(* IEC 61131-3 sources: POMIRTS_lab3/AS/Library_2/AsOpcUac, 3 files *)

(* ---- AsOpcUac.typ ---- *)
 TYPE
	UASecurityMsgMode :
	(												(* Message security modes *)
    	UASecurityMsgMode_BestAvailable 	:= 0,	(* Detects best available mode the server provides (may result in no security) 	*)
	  	UASecurityMsgMode_None          	:= 1,	(* No secure communication 														*)
	  	UASecurityMsgMode_Sign          	:= 2,	(* Messages are signed to verify peer authenticity 								*)
	  	UASecurityMsgMode_SignEncrypt   	:= 3	(* Messages are signed and encrypted 											*)
	);

  	UASecurityPolicy :
  	(												(* Security policies *)
    	UASecurityPolicy_BestAvailable  	:= 0,	(* Detects best available policy the server provides (may result in no security)	*)
    	UASecurityPolicy_None           	:= 1,	(* No secure communication (Allowed only for security mode = none)					*)
    	UASecurityPolicy_Basic128Rsa15  	:= 2,	(* RSA-PKCS-#1-V1.5-SHA1/RSA-PKCS-#1-V1.5/128-512 bit, HMAC-SHA1/AES-128-CBC/16bit	*)
    	UASecurityPolicy_Basic256       	:= 3,	(* RSA-PKCS-#1-OAEP-SHA1/RSA-OAEP/128-512 bit, HMAC-SHA1/AES-256-CBC/32bit			*)
    	UASecurityPolicy_Basic256Sha256   	:= 4	(* RSA-PKCS-#1-OAEP-SHA1/RSA-OAEP/256-512 bit, HMAC-SHA1/AES-256-CBC/32bit			*)
  	);

  	UATransportProfile :
  	(  												(* Transport profiles to select encoding and protocol *)
    	UATP_UATcp             				:= 1,	(* UA Binary over TCP								*)
    	UATP_WSHttpBinary      				:= 2,	(* Binary over HTTP			Not supported by B&R	*)
    	UATP_WSHttpXmlOrBinary 				:= 3,	(* XML/Binary over HTTP		Not supported by B&R	*)
    	UATP_WSHttpXml         				:= 4	(* XML over HTTP			Not supported by B&R	*)
  	);

 	UAUserIdentityTokenTtype :
 	(  												(* Authentication token type provided for logon *)
 		UAUITT_Anonymous					:= 0,	(* Logon anonymously					*)
 		UAUITT_Username						:= 1,	(* Logon with user name and password 	*)
 		UAUITT_x509							:= 2	(* Logon with user certificate			*)
 	);

	UAIdentifierType :
	(												(* Node identifier type *)
		UAIdentifierType_String 			:= 1,	(* String			*)
		UAIdentifierType_Numeric 			:= 2,	(* Numeric value	*)
		UAIdentifierType_GUID 				:= 3,	(* GUID				*)
		UAIdentifierType_Opaque				:= 4	(* ByteString		*)
	);

	UADeadbandType :
	(												(* Deadband type for monitored item sampling *)
		UADeadbandType_None 				:= 0,	(* No deadband, each value change is sampled						*)
		UADeadbandType_Absolute 			:= 1,	(* Absolute value to exceed from last sample to make new sample		*)
		UADeadbandType_Percent				:= 2	(* Percent of EURange to exceed from last sample to make new sample	*)
	);

	UANodeClass :
	(												(* Node classes defined through the OPC-UA standard *)
		UANodeClass_None 					:= 0,
		UANodeClass_Object					:= 1,
		UANodeClass_Variable 				:= 2,
		UANodeClass_Method					:= 4,
		UANodeClass_ObjectType				:= 8,
		UANodeClass_VariableType			:= 16,
		UANodeClass_ReferenceType			:= 32,
		UANodeClass_DataType				:= 64,
		UANodeClass_View					:= 128,
		UANodeClass_All						:= 255
	);

	UAAttributeId :
	(												(* Attributes defined through the OPC-UA standard *)
	  	UAAI_Default						:= 0,
		UAAI_NodeId							:= 1,
		UAAI_NodeClass						:= 2,
		UAAI_BrowseName						:= 3,
		UAAI_DisplayName					:= 4,
		UAAI_Description					:= 5,
		UAAI_WriteMask						:= 6,
		UAAI_UserWriteMask					:= 7,
		UAAI_IsAbstract						:= 8,
		UAAI_Symmetric						:= 9,
		UAAI_InverseName					:= 10,
		UAAI_ContainsNoLoops				:= 11,
		UAAI_EventNotifier					:= 12,
		UAAI_Value							:= 13,
		UAAI_DataType						:= 14,
		UAAI_ValueRank						:= 15,
		UAAI_ArrayDimensions				:= 16,
		UAAI_AccessLevel					:= 17,
		UAAI_UserAccessLevel				:= 18,
		UAAI_MinimumSamplingInterval		:= 19,
		UAAI_Historizing					:= 20,
		UAAI_Executable						:= 21,
		UAAI_UserExecutable					:= 22
	);

	UAConnectionStatus :
	(												(* Status of the underlying connection		*)
		UACS_Connected						:= 0,
		UACS_ConnectionError				:= 1,
		UACS_Shutdown						:= 2
	);

	UAServerState :
	(												(* State of the server read from Object.Server.ServerStatus.State	*)
		UASS_Running						:= 0,
		UASS_Failed							:= 1,
		UASS_NoConfiguration				:= 2,
		UASS_Suspended						:= 3,
		UASS_Shutdown						:= 4,
		UASS_Test							:= 5,
		UASS_CommunicationFault				:= 6,
		UASS_Unknown              			:= 7
	);

	UAVariantType :
	(												(* Kind of the variant data *)
		UAVariantType_Null					:= 0,	(* No data *)
		UAVariantType_Boolean				:= 1,	(* Data in element Boolean *)
		UAVariantType_SByte					:= 2,	(* Data in element SByte *)
		UAVariantType_Byte					:= 3,	(* Data in element Byte *)
		UAVariantType_Int16					:= 4,	(* Data in element Int16 *)
		UAVariantType_UInt16				:= 5,	(* Data in element UInt16 *)
		UAVariantType_Int32					:= 6,	(* Data in element Int32 *)
		UAVariantType_UInt32				:= 7,	(* Data in element UInt32 *)
		UAVariantType_Int64					:= 8,	(* Data in element Int64 *)
		UAVariantType_UInt64				:= 9,	(* Data in element UInt64 *)
		UAVariantType_Float					:= 10,	(* Data in element Float *)
		UAVariantType_Double				:= 11,	(* Data in element Double *)
		UAVariantType_String				:= 12,	(* Data in element String *)
		UAVariantType_DateTime				:= 13,	(* Data in element DateTime *)
		UAVariantType_Guid					:= 14,	(* Guid data in element String *)
		UAVariantType_ByteString			:= 15,	(* Byte string in element String *)
		UAVariantType_XmlElement			:= 16,	(* XML data in element String *)
		UAVariantType_NodeId				:= 17,	(* Data in element NodeId *)
		UAVariantType_ExpandedNodeId		:= 18,	(* Data in element ExpandedNodeId *)
		UAVariantType_StatusCode			:= 19,	(* Status code in element UInt32 *)
		UAVariantType_QualifiedName			:= 20,	(* Data in element QualifiedName *)
		UAVariantType_LocalizedText			:= 21	(* Data in element LocalizedText *)
	);

	UAArrayLength : DINT;							(* Arraylength of value attribute in AttributeRead and AttributeWrite services *)

	UANoOfElements : DINT;							(* Number of elements for arrays nested in structures *)

   	UAUserIdentityToken : STRUCT 					(* Identity token for authentication on an OPC-UA server *)
		UserIdentityTokenType	: UAUserIdentityTokenTtype;
		TokenParam1 			: STRING[255];
		TokenParam2				: STRING[255];
	END_STRUCT;

 	UASessionConnectInfo : STRUCT 					(* Session information and parameters *)
 	  	SessionName   			: STRING[255];
 	  	ApplicationName   		: STRING[255];
 	  	SecurityMsgMode   		: UASecurityMsgMode;
    	SecurityPolicy   		: UASecurityPolicy;
		CertificateStore		: STRING[255];
		ClientCertificateName	: STRING[255];
		ServerUri				: STRING[255];
		CheckServerCertificate	: BOOL;
    	TransportProfile 		: UATransportProfile;
    	UserIdentityToken		: UAUserIdentityToken;
		VendorSpecificParameter	: STRING[255];
    	SessionTimeout   		: TIME;
    	MonitorConnection		: TIME;
    	LocaleIDs				: ARRAY[0..4] OF STRING[6];
	END_STRUCT;

  	UANodeID : STRUCT 											(* Node identifier used to address nodes on the server		*)
		NamespaceIndex			: UINT;							(* Index of the namespace which contains the node			*)
		Identifier 				: STRING[255];					(* Node identifier according to the identifier types format *)
		IdentifierType			: UAIdentifierType; 			(* String, Numeric, GUID, ByteString						*)
	END_STRUCT;

	UAMonitoringSettings : STRUCT								(* Settings for data item monitoring						*)
		SamplingInterval		: TIME;							(* Time in ms 												*)
		DeadbandType			: UADeadbandType; 				(* Deadband type which applies to deadband value			*)
		Deadband				: REAL; 						(* Deadband value, semantics depending on DeadbandType 		*)
	END_STRUCT;

	UAMonitoringParameters : STRUCT								(* Settings for data item monitoring								*)
		SamplingInterval		: TIME;							(* Time in ms 														*)
		QueueSize				: UINT;							(* Size of the server sided queue to collect value changes			*)
		DiscardOldest			: BOOL;							(* True to discard oldest on queue overflow or newest otherwise		*)
		DeadbandType			: UADeadbandType; 				(* Deadband type which applies to deadband value					*)
		Deadband				: REAL; 						(* Deadband value, semantics depending on DeadbandType 				*)
	END_STRUCT;

	UALocalizedText : STRUCT									(* Localized text with locale identifer and text		*)
		Locale					: STRING[6];
		Text					: STRING[255];
	END_STRUCT;

	UANodeInfo : STRUCT											(* Node attribute values		*)
		AccessLevel 			: BYTE;
		ArrayDimension			: ARRAY[0..MAX_INDEX_ARRAYDIMENSION] OF UDINT;
		BrowseName				: STRING[255];
		ContainsNoLoops 		: BOOL;
		DataType				: UANodeID;
		Description				: UALocalizedText;
		DisplayName				: UALocalizedText;
		EventNotifier			: BYTE;
		Executable				: BOOL;
		Historizing				: BOOL;
		InverseName				: STRING[255];
		IsAbstract				: BOOL;
		MinimumSamplingInterval	: TIME;
		NodeClass				: UANodeClass;
		NodeID					: UANodeID;
		Symmetric				: BOOL;
		UserAccessLevel			: BYTE;
		UserExecutable			: BOOL;
		UserWriteMask			: UDINT;
		ValueRank				: DINT;
		WriteMask				: UDINT;
	END_STRUCT;

	UAIndexRange : STRUCT										(* Index range used for indexed access on arrays	*)
		StartIndex				: UINT;
		EndIndex 				: UINT;
	END_STRUCT;

	UANodeAdditionalInfo : STRUCT								(* Additional info for reading and writing node attributes	*)
		AttributeId				: UAAttributeId;
		IndexRangeCount			: UINT;
		IndexRange 				: ARRAY[0..MAX_INDEX_INDEXRANGE] OF UAIndexRange;
	END_STRUCT;

	UAMethodArgument : STRUCT						(* Method argument used to supply the input and receive the output argument values for method calls *)
		Name					: STRING[64];		(* Name of the method argument																		*)
		Value					: STRING[255];		(* Source/Destination variable name for the argument value											*)
	END_STRUCT;

	UAByteString : STRUCT							(* Byte string containing length and data	*)
		Length					: DINT;
		Data					: ARRAY[0..MAX_INDEX_BYTESTRING] OF USINT;
	END_STRUCT;

	UAExpandedNodeID : STRUCT 						(* Expanded node identfier type *)
		NodeId					: UANodeID;
		NamespaceUri			: STRING[255];
		ServerIndex				: UDINT;
	END_STRUCT;

	UAQualifiedName : STRUCT						(* Qualified name type *)
		NamespaceIndex			: UINT;
		Name					: STRING[255];
	END_STRUCT;

	UARelativePathElement : STRUCT					(* Relative path element used to build a relative path	*)
	    ReferenceTypeId			: UANodeID;
		IsInverse				: BOOL;
		IncludeSubTypes			: BOOL;
		TargetName				: UAQualifiedName;
	END_STRUCT;

	UARelativePath : STRUCT							(* Relative path used to translate and browse nodes	*)
	    NoOfElements			: DWORD;
		Elements				: ARRAY[0..MAX_INDEX_RELATIVEPATH] OF UARelativePathElement;
	END_STRUCT;

	UADataValue : STRUCT							(* Additional informations about data value *)
		Valid 					: BOOL;
		Reserved				: ARRAY[0..2]OF USINT;
		StatusCode				: UDINT;
		SourceTimestamp			: DATE_AND_TIME;
		ServerTimestamp			: DATE_AND_TIME;
	END_STRUCT;

	UAVariantData : STRUCT							(* Standard type for variant data *)
		VariantType				: UAVariantType;
		Boolean					: BOOL;
		SByte					: SINT;
		Byte					: USINT;
		Int16					: INT;
		UInt16					: UINT;
		Int32					: DINT;
		UInt32					: UDINT;
		Float					: REAL;
		Double					: LREAL;
		DateTime				: DATE_AND_TIME;
		String					: STRING[255];
		NodeId					: UANodeID;
		ExpandedNodeId			: UAExpandedNodeID;
		QualifiedName			: UAQualifiedName;
		LocalizedText			: UALocalizedText;
		DataValue				: UADataValue;
	END_STRUCT;

	UARange : STRUCT								(* Range for a value *)
		Low						: LREAL;
		High					: LREAL;
	END_STRUCT;

	UAEUInformation : STRUCT 						(* Information about the engineering units *)
		NamespaceUri			: STRING[255];
		UnitId					: DINT;
		DisplayName				: UALocalizedText;
		Description				: UALocalizedText;
	END_STRUCT;

	UATimeZoneData : STRUCT							(* Information about time zone	*)
		TimeOffset				: INT;				(* Offset in minutes from UTC	*)
		DaylightSaving			: BOOL;				(* Offset includes the DST		*)
	END_STRUCT;

	BrUaNodeId					: UANodeID;
	BrUaQualifiedName			: UAQualifiedName;
	BrUaLocalizedText			: UALocalizedText;
	BrUaByteString				: UAByteString;
	BrUaGuidString				: STRING[36];

	BrUaXmlElement : STRUCT
		Length					: DINT;
		Data					: STRING[65535];
	END_STRUCT;

	BrUaImageBMP : STRUCT
		Length					: DINT;
		Data					: ARRAY[0..6291455] OF USINT;
	END_STRUCT;
	BrUaImageGIF : STRUCT
		Length					: DINT;
		Data					: ARRAY[0..524287] OF USINT;
	END_STRUCT;
	BrUaImageJPG : STRUCT
		Length					: DINT;
		Data					: ARRAY[0..1048575] OF USINT;
	END_STRUCT;
	BrUaImagePNG : STRUCT
		Length					: DINT;
		Data					: ARRAY[0..2621439] OF USINT;
	END_STRUCT;

	BrUaDuration				: LREAL;
	BrUaLocaleIdString			: STRING[6];

	BrUaTimeZoneDataType		: UATimeZoneData;

END_TYPE

(* ---- AsOpcUac.fun ---- *)
{REDUND_CONTEXT} {REDUND_UNREPLICABLE} FUNCTION_BLOCK UA_Connect
	VAR_INPUT
		Execute	           		: BOOL;
		ServerEndpointUrl		: STRING[255];
		SessionConnectInfo 		: UASessionConnectInfo;
		Timeout            		: TIME;
	END_VAR

	VAR_OUTPUT
		ConnectionHdl      		: DWORD;
		Done			   		: BOOL;
		Busy               		: BOOL;
		Error              		: BOOL;
		ErrorID            		: DWORD;
	END_VAR

	VAR
		i_busy             		: BOOL;
	END_VAR
END_FUNCTION_BLOCK

{REDUND_CONTEXT} {REDUND_UNREPLICABLE} FUNCTION_BLOCK UA_Disconnect
	VAR_INPUT
		Execute	           		: BOOL;
		ConnectionHdl      		: DWORD;
		Timeout            		: TIME;
	END_VAR

	VAR_OUTPUT
		Done			   		: BOOL;
		Busy               		: BOOL;
		Error              		: BOOL;
		ErrorID            		: DWORD;
	END_VAR

	VAR
		i_busy             		: BOOL;
	END_VAR
END_FUNCTION_BLOCK

{REDUND_CONTEXT} {REDUND_UNREPLICABLE} FUNCTION_BLOCK UA_GetNamespaceIndex
	VAR_INPUT
		Execute	           		: BOOL;
		ConnectionHdl      		: DWORD;
		NamespaceUri			: STRING[255];
		Timeout            		: TIME;
	END_VAR

	VAR_OUTPUT
		NamespaceIndex			: UINT;
		Done			   		: BOOL;
		Busy               		: BOOL;
		Error              		: BOOL;
		ErrorID            		: DWORD;
	END_VAR

	VAR
		i_busy             		: BOOL;
	END_VAR
END_FUNCTION_BLOCK

{REDUND_CONTEXT} {REDUND_UNREPLICABLE} FUNCTION_BLOCK UA_TranslatePath
	VAR_INPUT
		Execute	           		: BOOL;
		ConnectionHdl      		: DWORD;
		StartNodeID				: UANodeID;
		RelativePath			: STRING[255];
		Timeout            		: TIME;
	END_VAR

	VAR_OUTPUT
		TargetNodeID			: UANodeID;
		Done			   		: BOOL;
		Busy               		: BOOL;
		Error              		: BOOL;
		ErrorID            		: DWORD;
	END_VAR

	VAR
		i_busy             		: BOOL;
	END_VAR
END_FUNCTION_BLOCK

{REDUND_CONTEXT} {REDUND_UNREPLICABLE} FUNCTION_BLOCK UA_NodeGetHandle
	VAR_INPUT
		Execute	           	 	: BOOL;
		ConnectionHdl      	 	: DWORD;
		NodeID					: UANodeID;
		Timeout            		: TIME;
	END_VAR

	VAR_OUTPUT
		NodeHdl					: DWORD;
		Done			   		: BOOL;
		Busy               		: BOOL;
		Error              		: BOOL;
		ErrorID            		: DWORD;
	END_VAR

	VAR
		i_busy             		: BOOL;
	END_VAR
END_FUNCTION_BLOCK

{REDUND_CONTEXT} {REDUND_UNREPLICABLE} FUNCTION_BLOCK UA_NodeGetHandleList
	VAR_INPUT
		Execute	           	 	: BOOL;
		ConnectionHdl      	 	: DWORD;
		NodeIDCount				: UINT;
		NodeIDs					: ARRAY[0..MAX_INDEX_NODELIST] OF UANodeID;
		Timeout            		: TIME;
	END_VAR

	VAR_OUTPUT
		NodeHdls				: ARRAY[0..MAX_INDEX_NODELIST] OF DWORD;
		Done			   		: BOOL;
		Busy               		: BOOL;
		Error              		: BOOL;
		ErrorID					: DWORD;
		NodeErrorIDs           	: ARRAY[0..MAX_INDEX_NODELIST] OF DWORD;
	END_VAR

	VAR
		i_busy             		: BOOL;
	END_VAR
END_FUNCTION_BLOCK

{REDUND_CONTEXT} {REDUND_UNREPLICABLE} FUNCTION_BLOCK UA_NodeReleaseHandle
	VAR_INPUT
		Execute	           		: BOOL;
		ConnectionHdl      		: DWORD;
		NodeHdl      	 		: DWORD;
		Timeout            		: TIME;
	END_VAR

	VAR_OUTPUT
		Done			   		: BOOL;
		Busy               		: BOOL;
		Error              		: BOOL;
		ErrorID            		: DWORD;
	END_VAR

	VAR
		i_busy             		: BOOL;
	END_VAR
END_FUNCTION_BLOCK

{REDUND_CONTEXT} {REDUND_UNREPLICABLE} FUNCTION_BLOCK UA_NodeReleaseHandleList
	VAR_INPUT
		Execute	           		: BOOL;
		ConnectionHdl      		: DWORD;
		NodeHdlCount   	 		: UINT;
		NodeHdls				: ARRAY[0..MAX_INDEX_NODELIST] OF DWORD;
		Timeout            		: TIME;
	END_VAR

	VAR_OUTPUT
		Done			   		: BOOL;
		Busy               		: BOOL;
		Error              		: BOOL;
		ErrorID					: DWORD;
		NodeErrorIDs           	: ARRAY[0..MAX_INDEX_NODELIST] OF DWORD;
	END_VAR

	VAR
		i_busy             		: BOOL;
	END_VAR
END_FUNCTION_BLOCK

{REDUND_CONTEXT} {REDUND_UNREPLICABLE} FUNCTION_BLOCK UA_NodeGetInfo
	VAR_INPUT
		Execute	           		: BOOL;
		ConnectionHdl      		: DWORD;
		NodeID					: UANodeID;
		Timeout            		: TIME;
	END_VAR

	VAR_OUTPUT
		NodeInfo				: UANodeInfo;
		Done			   		: BOOL;
		Busy               		: BOOL;
		Error              		: BOOL;
		ErrorID            		: DWORD;
	END_VAR

	VAR
		i_busy             		: BOOL;
	END_VAR
END_FUNCTION_BLOCK

{REDUND_CONTEXT} {REDUND_UNREPLICABLE} FUNCTION_BLOCK UA_SubscriptionCreate
	VAR_INPUT
		Execute	           		: BOOL;
		ConnectionHdl      		: DWORD;
		PublishingEnable		: BOOL;
		Priority				: BYTE;
		Timeout            		: TIME;
	END_VAR

	VAR_OUTPUT
		SubscriptionHdl			: DWORD;
		Done			   		: BOOL;
		Busy               		: BOOL;
		Error              		: BOOL;
		ErrorID            		: DWORD;
	END_VAR

	VAR_IN_OUT
		PublishingInterval		: TIME;
	END_VAR

	VAR
		i_busy             		: BOOL;
	END_VAR
END_FUNCTION_BLOCK

{REDUND_CONTEXT} {REDUND_UNREPLICABLE} FUNCTION_BLOCK UA_SubscriptionDelete
	VAR_INPUT
		Execute	           		: BOOL;
		SubscriptionHdl			: DWORD;
		Timeout            		: TIME;
	END_VAR

	VAR_OUTPUT
		Done			   		: BOOL;
		Busy               		: BOOL;
		Error              		: BOOL;
		ErrorID            		: DWORD;
	END_VAR

	VAR
		i_busy             		: BOOL;
	END_VAR
END_FUNCTION_BLOCK

{REDUND_CONTEXT} {REDUND_UNREPLICABLE} FUNCTION_BLOCK UA_SubscriptionOperate
	VAR_INPUT
		Execute	           		: BOOL;
		SubscriptionHdl			: DWORD;
		PublishingEnable  		: BOOL;
		Priority  				: USINT;
		Timeout            		: TIME;
	END_VAR

	VAR_OUTPUT
		Published				: BOOL;
		Done			   		: BOOL;
		Busy               		: BOOL;
		Error              		: BOOL;
		ErrorID            		: DWORD;
	END_VAR

	VAR_IN_OUT
		PublishingInterval		: TIME;
	END_VAR

	VAR
		i_busy             		: BOOL;
	END_VAR
END_FUNCTION_BLOCK

{REDUND_CONTEXT} {REDUND_UNREPLICABLE} FUNCTION_BLOCK UA_MonitoredItemAdd
	VAR_INPUT
		Execute	           		: BOOL;
		SubscriptionHdl			: DWORD;
		NodeHdl					: DWORD;
		NodeAddInfo				: UANodeAdditionalInfo;
		Timeout            		: TIME;
	END_VAR

	VAR_OUTPUT
		MonitoredItemHdl		: DWORD;
		Done			   		: BOOL;
		Busy               		: BOOL;
		Error              		: BOOL;
		ErrorID            		: DWORD;
	END_VAR

	VAR_IN_OUT
		Variable	   			: STRING[255];
		MonitoringSettings		: UAMonitoringSettings;
	END_VAR

	VAR
		i_busy             		: BOOL;
		i_tid					: UDINT;
	END_VAR
END_FUNCTION_BLOCK

{REDUND_CONTEXT} {REDUND_UNREPLICABLE} FUNCTION_BLOCK UA_MonitoredItemAddList
	VAR_INPUT
		Execute	           		: BOOL;
		SubscriptionHdl			: DWORD;
		NodeHdlCount			: UINT;
		NodeHdls				: ARRAY[0..MAX_INDEX_MONITORLIST] OF DWORD;
		NodeAddInfos			: ARRAY[0..MAX_INDEX_MONITORLIST] OF UANodeAdditionalInfo;
		Timeout            		: TIME;
	END_VAR

	VAR_OUTPUT
		Done			   		: BOOL;
		Busy               		: BOOL;
		Error              		: BOOL;
		ErrorID            		: DWORD;
		NodeErrorIDs			: ARRAY[0..MAX_INDEX_MONITORLIST] OF DWORD;
		MonitoredItemHdls		: ARRAY[0..MAX_INDEX_MONITORLIST] OF DWORD;
	END_VAR

	VAR_IN_OUT
		Variables	   			: ARRAY[0..MAX_INDEX_MONITORLIST] OF STRING[255];
		MonitoringSettings		: ARRAY[0..MAX_INDEX_MONITORLIST] OF UAMonitoringParameters;
		ValuesChanged			: ARRAY[0..MAX_INDEX_MONITORLIST] OF BOOL;
		RemainingValueCount		: ARRAY[0..MAX_INDEX_MONITORLIST] OF UINT;
		TimeStamps				: ARRAY[0..MAX_INDEX_MONITORLIST] OF DT;
		NodeQualityIDs			: ARRAY[0..MAX_INDEX_MONITORLIST] OF DWORD;
	END_VAR

	VAR
		i_busy             		: BOOL;
		i_tid					: UDINT;
	END_VAR
END_FUNCTION_BLOCK

{REDUND_CONTEXT} {REDUND_UNREPLICABLE} FUNCTION_BLOCK UA_MonitoredItemRemove
	VAR_INPUT
		Execute	           		: BOOL;
		MonitoredItemHdl		: DWORD;
		Timeout            		: TIME;
	END_VAR

	VAR_OUTPUT
		Done			   		: BOOL;
		Busy               		: BOOL;
		Error              		: BOOL;
		ErrorID            		: DWORD;
	END_VAR

	VAR
		i_busy             		: BOOL;
	END_VAR
END_FUNCTION_BLOCK

{REDUND_CONTEXT} {REDUND_UNREPLICABLE} FUNCTION_BLOCK UA_MonitoredItemRemoveList
	VAR_INPUT
		Execute	           		: BOOL;
		SubscriptionHdl			: DWORD;
		MonitoredItemHdlCount	: UINT;
		MonitoredItemHdls		: ARRAY[0..MAX_INDEX_MONITORLIST] OF DWORD;
		Timeout            		: TIME;
	END_VAR

	VAR_OUTPUT
		Done			   		: BOOL;
		Busy               		: BOOL;
		Error              		: BOOL;
		ErrorID            		: DWORD;
		NodeErrorIDs			: ARRAY[0..MAX_INDEX_MONITORLIST] OF DWORD;
	END_VAR

	VAR
		i_busy             		: BOOL;
	END_VAR
END_FUNCTION_BLOCK

{REDUND_CONTEXT} {REDUND_UNREPLICABLE} FUNCTION_BLOCK UA_MonitoredItemOperate
	VAR_INPUT
		Execute	           		: BOOL;
		MonitoredItemHdl		: DWORD;
		Timeout            		: TIME;
	END_VAR

	VAR_OUTPUT
		ValueChanged			: BOOL;
		TimeStamp				: DT;
		Done			   		: BOOL;
		Busy               		: BOOL;
		Error              		: BOOL;
		ErrorID            		: DWORD;
	END_VAR

	VAR_IN_OUT
		MonitoringSettings 		: UAMonitoringSettings;
	END_VAR

	VAR
		i_busy             		: BOOL;
	END_VAR
END_FUNCTION_BLOCK

{REDUND_CONTEXT} {REDUND_UNREPLICABLE} FUNCTION_BLOCK UA_MonitoredItemOperateList
	VAR_INPUT
		Execute	           		: BOOL;
		SubscriptionHdl			: DWORD;
		MonitoredItemHdlCount	: UINT;
		MonitoredItemHdls		: ARRAY[0..MAX_INDEX_MONITORLIST] OF DWORD;
	END_VAR

	VAR_OUTPUT
		Published				: BOOL;
		Done			   		: BOOL;
		Busy               		: BOOL;
		Error              		: BOOL;
		ErrorID            		: DWORD;
		NodeErrorIDs			: ARRAY[0..MAX_INDEX_MONITORLIST] OF DWORD;
	END_VAR

	VAR
		i_busy             		: BOOL;
	END_VAR
END_FUNCTION_BLOCK

{REDUND_CONTEXT} {REDUND_UNREPLICABLE} FUNCTION_BLOCK UA_EventItemAdd
	VAR_INPUT
		Execute	           		: BOOL;
		SubscriptionHdl			: DWORD;
		NodeHdl					: DWORD;
		EventType				: UANodeID;
		EventFieldSelectionCount: UINT;
		EventFieldSelections	: ARRAY[0..MAX_INDEX_EVENTFIELDSELECTION] OF UARelativePath;
		Timeout            		: TIME;
	END_VAR

	VAR_OUTPUT
		EventItemHdl			: DWORD;
		Done			   		: BOOL;
		Busy               		: BOOL;
		Error              		: BOOL;
		ErrorID            		: DWORD;
	END_VAR

	VAR_IN_OUT
		EventFields	   			: ARRAY[0..MAX_INDEX_EVENTFIELDSELECTION] OF STRING[MAX_LENGTH_VARIABLE];
	END_VAR

	VAR
		i_busy             		: BOOL;
		i_tid					: UDINT;
	END_VAR
END_FUNCTION_BLOCK

{REDUND_CONTEXT} {REDUND_UNREPLICABLE} FUNCTION_BLOCK UA_EventItemRemove
	VAR_INPUT
		Execute	           		: BOOL;
		SubscriptionHdl			: DWORD;
		EventItemHdl			: DWORD;
		Timeout            		: TIME;
	END_VAR

	VAR_OUTPUT
		Done			   		: BOOL;
		Busy               		: BOOL;
		Error              		: BOOL;
		ErrorID            		: DWORD;
	END_VAR

	VAR
		i_busy             		: BOOL;
		i_tid					: UDINT;
	END_VAR
END_FUNCTION_BLOCK

{REDUND_CONTEXT} {REDUND_UNREPLICABLE} FUNCTION_BLOCK UA_EventItemOperate
	VAR_INPUT
		Execute	           		: BOOL;
		SubscriptionHdl			: DWORD;
		EventItemHdl			: DWORD;
		Timeout            		: TIME;
	END_VAR

	VAR_OUTPUT
		EventProcessed			: BOOL;
		RemainingEventCount		: INT;
		FieldErrorIDs			: ARRAY[0..MAX_INDEX_EVENTFIELDSELECTION] OF DWORD;
		Done			   		: BOOL;
		Busy               		: BOOL;
		Error              		: BOOL;
		ErrorID            		: DWORD;
	END_VAR

	VAR
		i_busy             		: BOOL;
		i_tid					: UDINT;
	END_VAR
END_FUNCTION_BLOCK

{REDUND_CONTEXT} {REDUND_UNREPLICABLE} FUNCTION_BLOCK UA_Read
	VAR_INPUT
		Execute	           		: BOOL;
		ConnectionHdl      		: DWORD;
		NodeHdl					: DWORD;
		NodeAddInfo				: UANodeAdditionalInfo;
		Timeout            		: TIME;
	END_VAR

	VAR_OUTPUT
		Done			   		: BOOL;
		Busy               		: BOOL;
		Error              		: BOOL;
		ErrorID            		: DWORD;
		TimeStamp				: DT;
	END_VAR

	VAR_IN_OUT
		Variable	   			: STRING[255];
	END_VAR

	VAR
		i_busy             		: BOOL;
		i_tid					: UDINT;
	END_VAR
END_FUNCTION_BLOCK

{REDUND_CONTEXT} {REDUND_UNREPLICABLE} FUNCTION_BLOCK UA_ReadList
	VAR_INPUT
		Execute	           		: BOOL;
		ConnectionHdl      		: DWORD;
		NodeHdlCount			: UINT;
		NodeHdls				: ARRAY[0..MAX_INDEX_NODELIST] OF DWORD;
		NodeAddInfo				: ARRAY[0..MAX_INDEX_NODELIST] OF UANodeAdditionalInfo;
		Timeout            		: TIME;
	END_VAR

	VAR_OUTPUT
		Done			   		: BOOL;
		Busy               		: BOOL;
		Error              		: BOOL;
		ErrorID            		: DWORD;
		NodeErrorIDs			: ARRAY[0..MAX_INDEX_NODELIST] OF DWORD;
		TimeStamps				: ARRAY[0..MAX_INDEX_NODELIST] OF DT;
	END_VAR

	VAR_IN_OUT
		Variables	   			: ARRAY[0..MAX_INDEX_NODELIST] OF STRING[255];
	END_VAR

	VAR
		i_busy             		: BOOL;
		i_tid					: UDINT;
	END_VAR
END_FUNCTION_BLOCK

{REDUND_CONTEXT} {REDUND_UNREPLICABLE} FUNCTION_BLOCK UaClt_ReadBulk
	VAR_INPUT
		Execute	           		: BOOL;
		ConnectionHdl      		: DWORD;
		NodeIDCount				: UINT;
		NodeIDs					: UDINT;
		NodeAddInfo				: UDINT;
		Variables	   			: UDINT;
		NodeErrorIDs			: UDINT;
		TimeStamps				: UDINT;
		Timeout            		: TIME;
	END_VAR

	VAR_OUTPUT
		Done			   		: BOOL;
		Busy               		: BOOL;
		Error              		: BOOL;
		ErrorID            		: DWORD;
	END_VAR

	VAR
		i_busy             		: BOOL;
		i_tid					: UDINT;
	END_VAR
END_FUNCTION_BLOCK

{REDUND_CONTEXT} {REDUND_UNREPLICABLE} FUNCTION_BLOCK UA_Write
	VAR_INPUT
		Execute	           		: BOOL;
		ConnectionHdl      		: DWORD;
		NodeHdl					: DWORD;
		NodeAddInfo				: UANodeAdditionalInfo;
		Timeout            		: TIME;
	END_VAR

	VAR_OUTPUT
		Done			   		: BOOL;
		Busy               		: BOOL;
		Error              		: BOOL;
		ErrorID            		: DWORD;
	END_VAR

	VAR_IN_OUT
		Variable	   			: STRING[255];
	END_VAR

	VAR
		i_busy             		: BOOL;
		i_tid					: UDINT;
	END_VAR
END_FUNCTION_BLOCK

{REDUND_CONTEXT} {REDUND_UNREPLICABLE} FUNCTION_BLOCK UA_WriteList
	VAR_INPUT
		Execute	           		: BOOL;
		ConnectionHdl      		: DWORD;
		NodeHdlCount			: UINT;
		NodeHdls				: ARRAY[0..MAX_INDEX_NODELIST] OF DWORD;
		NodeAddInfo				: ARRAY[0..MAX_INDEX_NODELIST] OF UANodeAdditionalInfo;
		Timeout            		: TIME;
	END_VAR

	VAR_OUTPUT
		Done			   		: BOOL;
		Busy               		: BOOL;
		Error              		: BOOL;
		ErrorID            		: DWORD;
		NodeErrorIDs			: ARRAY[0..MAX_INDEX_NODELIST] OF DWORD;
	END_VAR

	VAR_IN_OUT
		Variables   			: ARRAY[0..MAX_INDEX_NODELIST] OF STRING[255];
	END_VAR

	VAR
		i_busy             		: BOOL;
		i_tid					: UDINT;
	END_VAR
END_FUNCTION_BLOCK

{REDUND_CONTEXT} {REDUND_UNREPLICABLE} FUNCTION_BLOCK UaClt_WriteBulk
	VAR_INPUT
		Execute	           		: BOOL;
		ConnectionHdl      		: DWORD;
		NodeIDCount				: UINT;
		NodeIDs					: UDINT;
		NodeAddInfo				: UDINT;
		Variables	   			: UDINT;
		NodeErrorIDs			: UDINT;
		Timeout            		: TIME;
	END_VAR

	VAR_OUTPUT
		Done			   		: BOOL;
		Busy               		: BOOL;
		Error              		: BOOL;
		ErrorID            		: DWORD;
	END_VAR

	VAR
		i_busy             		: BOOL;
		i_tid					: UDINT;
	END_VAR
END_FUNCTION_BLOCK

{REDUND_CONTEXT} {REDUND_UNREPLICABLE} FUNCTION_BLOCK UA_MethodGetHandle
	VAR_INPUT
		Execute	           		: BOOL;
		ConnectionHdl      		: DWORD;
		ObjectNodeID			: UANodeID;
		MethodNodeID			: UANodeID;
		Timeout            		: TIME;
	END_VAR

	VAR_OUTPUT
		MethodHdl				: DWORD;
		Done			   		: BOOL;
		Busy               		: BOOL;
		Error              		: BOOL;
		ErrorID            		: DWORD;
	END_VAR

	VAR
		i_busy             		: BOOL;
	END_VAR
END_FUNCTION_BLOCK

{REDUND_CONTEXT} {REDUND_UNREPLICABLE} FUNCTION_BLOCK UA_MethodReleaseHandle
	VAR_INPUT
		Execute	           		: BOOL;
		ConnectionHdl      		: DWORD;
		MethodHdl				: DWORD;
		Timeout            		: TIME;
	END_VAR

	VAR_OUTPUT
		Done			   		: BOOL;
		Busy               		: BOOL;
		Error              		: BOOL;
		ErrorID            		: DWORD;
	END_VAR

	VAR
		i_busy             		: BOOL;
	END_VAR
END_FUNCTION_BLOCK

{REDUND_CONTEXT} {REDUND_UNREPLICABLE} FUNCTION_BLOCK UA_MethodCall
	VAR_INPUT
		Execute	           		: BOOL;
		ConnectionHdl      		: DWORD;
		MethodHdl				: DWORD;
		Timeout            		: TIME;
	END_VAR

	VAR_OUTPUT
		Done			   		: BOOL;
		Busy               		: BOOL;
		Error              		: BOOL;
		ErrorID            		: DWORD;
	END_VAR

	VAR_IN_OUT
		InputArguments			: ARRAY[0..MAX_INDEX_ARGUMENTS] OF UAMethodArgument;
		OutputArguments			: ARRAY[0..MAX_INDEX_ARGUMENTS] OF UAMethodArgument;
	END_VAR

	VAR
		i_busy             		: BOOL;
		i_tid					: UDINT;
	END_VAR
END_FUNCTION_BLOCK

{REDUND_CONTEXT} {REDUND_UNREPLICABLE} FUNCTION_BLOCK UA_ConnectionGetStatus
	VAR_INPUT
		Execute	           		: BOOL;
		ConnectionHdl      		: DWORD;
		Timeout            		: TIME;
	END_VAR

	VAR_OUTPUT
		ConnectionStatus		: UAConnectionStatus;
		ServerState				: UAServerState;
		ServiceLevel			: BYTE;
		Done			   		: BOOL;
		Busy               		: BOOL;
		Error              		: BOOL;
		ErrorID            		: DWORD;
	END_VAR

	VAR
		i_busy             		: BOOL;
	END_VAR
END_FUNCTION_BLOCK

(* ---- AsOpcUac.var ---- *)
VAR CONSTANT
	MAX_LENGTH_VARIABLE					: UINT := 255;
	MAX_LENGTH_BYTESTRING				: UINT := 1024;

	MAX_ELEMENTS_ARRAYDIMENSION 		: UINT := 7;	(* B&R supports arrays with 7 dimensions											*)
	MAX_ELEMENTS_INDEXRANGE 			: UINT := 8;	(* Index range addresses max number of dimensions +1 for string/bytestring index	*)
	MAX_ELEMENTS_NODELIST 				: UINT := 64;	(* Maximum number of items the node list functions can handle						*)
	MAX_ELEMENTS_MONITORLIST			: UINT := 64;	(* Maximum number of elements the monitored item list functions can handle			*)
	MAX_ELEMENTS_ARGUMENTS 				: UINT := 10;	(* Maximum number of input and output arguments for method call						*)
	MAX_ELEMENTS_EVENTFIELDSELECTION	: UINT := 64;
	MAX_ELEMENTS_RELATIVEPATH			: UINT := 16;

	(* B&R requires zero based arrays in .typ and .fun files, calculations like "const - 1" are not allowed
	   for declarations in those files, so other constants denoting the array upper limit are declared *)
	MAX_INDEX_ARRAYDIMENSION 			: UINT := MAX_ELEMENTS_ARRAYDIMENSION - 1;
	MAX_INDEX_INDEXRANGE 				: UINT := MAX_ELEMENTS_INDEXRANGE - 1;
	MAX_INDEX_NODELIST 					: UINT := MAX_ELEMENTS_NODELIST - 1;
	MAX_INDEX_MONITORLIST 				: UINT := MAX_ELEMENTS_MONITORLIST - 1;
	MAX_INDEX_ARGUMENTS 				: UINT := MAX_ELEMENTS_ARGUMENTS - 1;
	MAX_INDEX_EVENTFIELDSELECTION		: UINT := MAX_ELEMENTS_EVENTFIELDSELECTION - 1;
	MAX_INDEX_RELATIVEPATH				: UINT := MAX_ELEMENTS_RELATIVEPATH - 1;
	MAX_INDEX_BYTESTRING				: UINT := MAX_LENGTH_BYTESTRING - 1;
END_VAR
